(* IEC 61131-3 sources: tsplc/packages/build/tests/fixtures/raw-st/src, 1 file *)

(* ---- Main.st ---- *)
PROGRAM Main
VAR
	Station : FB_FillingStation;
END_VAR
PRG_ReadInputs();
PRG_Transport();
Station();
PRG_Publish();
END_PROGRAM
